TYPE ST_ControlValveStateMachineTest :
STRUCT
    calibrationTimerDone : BOOL;
    simulatedOpenElapsedTime : TIME;
    simulatedCloseElapsedTime : TIME;
	simulatedOpeningPercentage : DINT;
END_STRUCT
END_TYPE

(* stored: Version 1.1.0.1, ProductVersion 3.1.4024.9
   DUT ST_ControlValveStateMachineTest: Id {99c3b690-225c-4fb6-a66f-6aba732b46af} *)
